Fanuc KAREL source: KS00043.KL

PROGRAM KS00043
%NOLOCKGROUP
TYPE
  REC_T = STRUCTURE
    VALUE: INTEGER
    FLAG: BOOLEAN
  ENDSTRUCTURE
VAR
  A: ARRAY[4] OF XYZWPREXT
  B: ARRAY[4] OF XYZWPREXT
  FLAG: BOOLEAN
  N: INTEGER
  STATUS: INTEGER
  PN: STRING[80]
  VN: STRING[80]
BEGIN
  PN = ''
  VN = 'A'
  FLAG = A = B
END KS00043
